(* IEC 61131-3 sources: Test-Git_ESME26/TestProgettoESME_26.fbsproj/PacDriveLib_Motion_Migration_Example.device.xml.v3^/Plc Logic.plclogic.xml.v3^/Application.application.xml.v3^/Test_YOffset, 1 file *)

(* ---- SR_YOffset.prg.st ---- *)
PROGRAM SR_YOffset
VAR
	xInitDone					: BOOL;
	xInitError					: BOOL;
	etResult					: MOIN.ET_Result;

	fbDriveEnable				: PDL_FB_DriveEnable;
	fbYOffsetCorrection			: PDL_FB_YOffsetCorrection;
	fbVarioPosJerk				: PDL_FB_VarioPosJerk;
END_VAR

IF  NOT xInitDone
THEN

	IF  SR_Sercos.q_xSercosRun
	THEN
		xInitDone := TRUE;

		fbVarioPosJerk.i_lrAcc   		:= 1000;
		fbVarioPosJerk.i_lrDec  		:= 1000;
		fbVarioPosJerk.i_lrJerk 		:= 1000;
		fbVarioPosJerk.i_lrVel   		:= 100;
		fbVarioPosJerk.i_lrTarget 		:= 200;
		fbVarioPosJerk.i_etPosMode		:= PDL_ET_PosMode.Absolute;

		Logical_Encoder_YOffset.ConnectMasterAxis( i_ifAxis := DRV_YOffset.Axis,
													q_xError   => xInitError,
													q_etResult => etResult
													);

		fbYOffsetCorrection.i_lrCorrection 	:= 100;
		fbYOffsetCorrection.i_lrMaxCorrAcc 	:= 1000;
		fbYOffsetCorrection.i_lrMaxCorrVel 	:= 100;
		fbYOffsetCorrection.i_lrXFactor 	:= 50;
		fbYOffsetCorrection.i_lrXStartPos 	:= 100;
	END_IF
END_IF

fbDriveEnable( i_ifDrive := DRV_YOffset.Axis );

fbYOffsetCorrection( 	i_ifDrive 	 := DRV_YOffset.Axis,
						i_lencMaster := Logical_Encoder_YOffset );

//pos mode endless does not work with channel (setpos not working)
fbVarioPosJerk( i_ifDrive := fbYOffsetCorrection.ifGetControlChannel );
